(* IEC 61131-3 sources: Test002/ConveyorBelt/Class/SafetyBaseFSoE (part 4) *)

    // if searched path has been found, we already got this pdo in our list
    if (PdoCfg.SourcePathLen = pHelp^.PdoInfo.SourcePathLen) & (PdoCfg.DestPathLen = pHelp^.PdoInfo.DestPathLen) &
      (PdoCfg.InterfaceCRC = pHelp^.PdoInfo.InterfaceCRC) &
      (ToStdLib.MemCmp(dest:= PdoCfg.pSourcePath, source:= pHelp^.PdoInfo.pSourcePath , size:= PdoCfg.SourcePathLen) = 0) &
      (ToStdLib.MemCmp(dest:= PdoCfg.pDestPath,   source:= pHelp^.PdoInfo.pDestPath   , size:= PdoCfg.DestPathLen  ) = 0) then
      // already in buffer => leave function
      return;
    else
      pHelp^.pNext$pvoid := ToStdLib.Malloc(size:=sizeof(t_PdoListElem));
      pHelp := pHelp^.pNext;
    end_if;
  end_if;

  if pHelp <> NIL then
    // allocate memory for the module source path
    pHelp^.PdoInfo.pSourcePath$pVoid := ToStdLib.Malloc(size:=PdoCfg.SourcePathLen);
    if pHelp^.PdoInfo.pSourcePath = NIL then
      SetSafetyState(NewState:=_MemAllocFailed);
      retcode := -1;
      return;
    end_if;

    _memcpy(ptr1:=pHelp^.PdoInfo.pSourcePath, ptr2:=PdoCfg.pSourcePath, cntr:=PdoCfg.SourcePathLen);

    // allocate memory for the module source path
    pHelp^.PdoInfo.pDestPath$pVoid := ToStdLib.Malloc(size:=PdoCfg.DestPathLen);
    if pHelp^.PdoInfo.pDestPath = NIL then
      SetSafetyState(NewState:=_MemAllocFailed);
      retcode := -1;
      return;
    end_if;

    _memcpy(ptr1:=pHelp^.PdoInfo.pDestPath, ptr2:=PdoCfg.pDestPath, cntr:=PdoCfg.DestPathLen);

    pHelp^.PdoInfo.Info           := PdoCfg.Info;
    pHelp^.PdoInfo.InterfaceCRC   := PdoCfg.InterfaceCRC;
    pHelp^.PdoInfo.SourcePathLen  := PdoCfg.SourcePathLen;
    pHelp^.PdoInfo.DestPathLen    := PdoCfg.DestPathLen;
    // length is only zero for non-interface pdos
    if PdoCfg.Info.IsInterfacePDO = FALSE then
      pHelp^.PdoInfo.PdoLen       := 0;   // the length is determined later in method CreateAndSendCfg
    else
      pHelp^.PdoInfo.PdoLen       := PdoCfg.PdoLen;
    end_if;
    pHelp^.PdoInfo.PDO_ID         := 255; // the ID is assigned later by the safety manager of the master domain
    pHelp^.pNext                  := NIL;

    PdoCfgNo += 1;
  else
    SetSafetyState(NewState:=_MemAllocFailed);
    retcode := -1;
    return;
  end_if;

END_FUNCTION

FUNCTION VIRTUAL SafetyBaseFSoE::AddSlaveToCfg
  VAR_INPUT
    pModule 	: ^SafetyBaseFSoE::PathInfoType;
    b_IsOptional 	: BOOL;
    b_IsInterface 	: BOOL;(* := FALSE *)
    InterfaceCRC 	: HDINT;(* := 0 *)
  END_VAR
  VAR
    pHelp : ^t_SlaveListElem;
  END_VAR

  if pFirstSlaveCfg = NIL then
    pFirstSlaveCfg$pVoid := ToStdLib.Malloc(size:=sizeof(t_SlaveListElem));
    pHelp := pFirstSlaveCfg;
  else
    pHelp := pFirstSlaveCfg;
    while pHelp^.pNext <> NIL do
      //if searched path is found, we already got this module in our list
      if (pModule^.ui_PathCompLen = pHelp^.SlaveInfo.CompPathLen) &
        (ToStdLib.MemCmp(dest:= pModule^.p_us_PathComp, source:= pHelp^.SlaveInfo.pCompPath , size:= pModule^.ui_PathCompLen) = 0) then
        // already in buffer => leave function
        return;
      else
        pHelp := pHelp^.pNext;
      end_if;
    end_while;

    //if searched path is found, we already got this module in our list
    if (pModule^.ui_PathCompLen = pHelp^.SlaveInfo.CompPathLen) &
      (ToStdLib.MemCmp(dest:= pModule^.p_us_PathComp, source:= pHelp^.SlaveInfo.pCompPath , size:= pModule^.ui_PathCompLen) = 0) then
      // already in buffer => leave function
      return;
    end_if;

    pHelp^.pNext$pvoid := ToStdLib.Malloc(size:=sizeof(t_SlaveListElem));
    pHelp := pHelp^.pNext;
  end_if;

  if pHelp <> NIL then
    // allocate memory for the module path
    pHelp^.SlaveInfo.PathLen := pModule^.p_us_Path^$UINT + 2;
    pHelp^.SlaveInfo.pPath$pVoid := ToStdLib.Malloc(size:=pHelp^.SlaveInfo.PathLen);
    if pHelp^.SlaveInfo.pPath = NIL then
      SetSafetyState(NewState:=_MemAllocFailed);
      LogError("@0243 (SafetyBaseFSoE::AddSlaveToCfg) Error: Failed to allocate memory for the module path.");
      return;
    end_if;

    _memcpy(ptr1:=pHelp^.SlaveInfo.pPath, ptr2:=pModule^.p_us_Path, cntr:=pHelp^.SlaveInfo.PathLen);

    // allocate memory for the module path
    pHelp^.SlaveInfo.CompPathLen := pModule^.ui_PathCompLen;
    pHelp^.SlaveInfo.pCompPath$pVoid := ToStdLib.Malloc(size:=pHelp^.SlaveInfo.CompPathLen);
    if pHelp^.SlaveInfo.pCompPath = NIL then
      SetSafetyState(NewState:=_MemAllocFailed);
      LogError("@0244 (SafetyBaseFSoE::AddSlaveToCfg) Error: Failed to allocate memory for the compressed module path.");
      return;
    end_if;

    _memcpy(ptr1:=pHelp^.SlaveInfo.pCompPath, ptr2:=pModule^.p_us_PathComp, cntr:=pHelp^.SlaveInfo.CompPathLen);

    pHelp^.SlaveInfo.Info             := 0;
    pHelp^.SlaveInfo.Info.IsOptional  := b_IsOptional;
    pHelp^.SlaveInfo.Info.IsInterface := b_IsInterface;

    pHelp^.SlaveInfo.InterfaceCRC := InterfaceCRC;

    pHelp^.pNext                  := NIL;

    SlaveCfgNo += 1;
  else
    SetSafetyState(NewState:=_MemAllocFailed);
    LogError("@0243 (SafetyBaseFSoE::AddSlaveToCfg) Error: Failed to allocate memory for the new list-element.");
    return;
  end_if;

END_FUNCTION

FUNCTION VIRTUAL SafetyBaseFSoE::FreeCfgLists
  VAR
    pHelpModule : ^t_ModuleListElem;
    pHelpPdo : ^t_PdoListElem;
    pHelpSlave : ^t_SlaveListElem;
//    pHelpUnsafeVar : ^t_UnsafeVarListElem;
  END_VAR

  // while we got module cfgs
  while pFirstModuleCfg do
    pHelpModule := pFirstModuleCfg;
    pFirstModuleCfg := pFirstModuleCfg^.pNext;

    if pHelpModule^.ModuleInfo.pDestCRCs then
      ToStdLib.Free(pHelpModule^.ModuleInfo.pDestCRCs);
    end_if;
    ToStdLib.Free(pHelpModule^.ModuleInfo.pPath);
    ToStdLib.Free(pHelpModule^.ModuleInfo.pCompPath);
    ToStdLib.Free(pHelpModule);
  end_while;
  pFirstModuleCfg := NIL;
  ModuleCfgNo := 0;

  // while we got pdo cfgs
  while pFirstPdoCfg do
    pHelpPdo := pFirstPdoCfg;
    pFirstPdoCfg := pFirstPdoCfg^.pNext;

    ToStdLib.Free(pHelpPdo^.PdoInfo.pSourcePath);
    ToStdLib.Free(pHelpPdo^.PdoInfo.pDestPath);
    ToStdLib.Free(pHelpPdo);
  end_while;
  pFirstPdoCfg := NIL;
  PdoCfgNo := 0;

  // while we got slave cfgs
  while pFirstSlaveCfg do
    pHelpSlave := pFirstSlaveCfg;
    pFirstSlaveCfg := pFirstSlaveCfg^.pNext;

    ToStdLib.Free(pHelpSlave^.SlaveInfo.pPath);
    ToStdLib.Free(pHelpSlave^.SlaveInfo.pCompPath);
    ToStdLib.Free(pHelpSlave);
  end_while;
  pFirstSlaveCfg := NIL;
  SlaveCfgNo := 0;

  FreeFSoEConnectionInfos();

// memory is freed by safety manager
//  // while we got unsafevar cfgs
//  while pFirstUnsafeCfg do
//    pHelpUnsafeVar := pFirstUnsafeCfg;
//    pFirstUnsafeCfg := pFirstUnsafeCfg^.pNext;
//
//    ToStdLib.Free(pHelpUnsafeVar^.UnsafeVarInfo.pName);
//    ToStdLib.Free(pHelpUnsafeVar);
//  end_while;
//  pFirstUnsafeCfg := NIL;
//  UnsafeCfgNo := 0;

  // reduze size of config mem used to 4 (only safety number of cpu module)
  ConfigMemSizeUsed := 4;

END_FUNCTION

FUNCTION VIRTUAL SafetyBaseFSoE::CreateAndSendCfg
  VAR
    pHelpModule       : ^t_ModuleListElem;
    pHelpPdo          : ^t_PdoListElem;
    pHelpSlave        : ^t_SlaveListElem;
    pHelpConnection   : ^t_FSoEConnectionDetails;
    pCfg              : ^void;
    TmpPathLen        : UINT;
    MyPara 	          : CmdStruct;
    MyResult	        : results;
    AddConfigSize     : UDINT;
    i                 : UDINT;
  END_VAR

(*
    Memory structure:
      4 Byte: SafetyNumber of CPU (is already there from initialisation in CSCP011_IM::InitSafeModule)
      1 Byte: Number of module configurations which are following
      for every module configuration (first is always the CPU itself)
        1 Byte: Info
        4 Byte: Interface Frame Source SafetyNumber (0 if it is no source for interface frames)
        4 Byte: Interface Frame CRC
        1 Byte: Number of destination inferface frame CRCs
        x Byte: Destination interface frame CRCs (number * sizeof(HDINT)
        2 Byte: Length of hardware path
        x Byte (depending on length in the 2 byte before): Hardwarepath
        2 Byte: Length of compressed hardware path
        x Byte (depending on length in the 2 byte before): Compressed Hardwarepath
        1 Byte: PDO out length for this module
      1 Byte: Number of pdo configurations which are following
      for every PDO configuration
        1 Byte: PDO length
        1 Byte: Interface frame info
        4 Byte: Interface CRC
        2 Byte: Length of source hardware path
        x Byte (depending on length in the 2 byte before): Hardwarepath of source
        2 Byte: Length of destination hardware path
        x Byte (depending on length in the 2 byte before): Hardwarepath of destination
      1 Byte: Number of slave configurations which are following
      for every slave configuration
        1 Byte: Info
        4 Byte: InterfaceCRC
        2 Byte: Length of hardware path
        x Byte (depending on length in the 2 byte before): Hardwarepath
        2 Byte: Length of compressed hardware path
        x Byte (depending on length in the 2 byte before): Compressed Hardwarepath
      2 Byte: Number of connection infos which are following
      for every FSoE connection info
        2 Byte: ConnectionID
        1 Byte: ConnectionState
        1 Byte: Flags // Actually, type is 4 bytes in size but for compatibility reasons it is still used as 1 byte. As a result, bits 9-32 are currently not used.
        4 Byte: Master safety number

only if feature available:
        2 Byte: Transmission time in ms

        2 Byte: Offset where to read from master
        2 Byte: Size of data to read from master (and write to slave)
        2 Byte: Offset where to write to master
        2 Byte: Size of data to write to master (and read from slave)
        2 Byte: SlaveAddress
        2 Byte: Length of slave hardware path
        x Byte (depending on length in the 2 byte before): Slave hardware path
        2 Byte: Length of compressed slave hardware path
        x Byte (depending on length in the 2 byte before): Compressed slave hardware path
        2 Byte: Offset where to read from slave
        2 Byte: Offset where to write to slave
*)

  // check if there is memory and if the only thing inside is the safety number
  if pConfigMem & (ConfigMemSizeUsed = 4) then
    // insert the safety number
    pConfigMem^$UDINT := SafetyNumber;

    // pCfg points to the next memory we have to write to => set it to the memory after the safety number
    pCfg := pConfigMem + ConfigMemSizeUsed;

    // add all module configurations to memory
    if pFirstModuleCfg then
      // add number of module configurations to memory (no need to check the memory here, because already 512 bytes are allocated)
      pCfg^$USINT       := ModuleCfgNo;
      pCfg              += sizeof(USINT);
      ConfigMemSizeUsed += sizeof(USINT);

      pHelpModule := pFirstModuleCfg;
      // go through list
      while pHelpModule do
        // add the elements

        // check if we have enough memory to add the next module
        AddConfigSize := sizeof(BSINT) + sizeof(HDINT) + sizeof(HDINT) + sizeof(UINT) + pHelpModule^.ModuleInfo.PathLen + sizeof(UINT) + pHelpModule^.ModuleInfo.CompPathLen + sizeof(USINT);
        if pHelpModule^.ModuleInfo.Info.IsInterfaceDest then
          AddConfigSize += sizeof(USINT) + pHelpModule^.ModuleInfo.DestCRCNo * sizeof(HDINT);
        end_if;

        pCfg := CheckConfigMemSize(AddConfigSize);
        if pCfg = NIL then
          // error message already logged by function
          return;
        end_if;

        // info
        pCfg^$BSINT := pHelpModule^.ModuleInfo.Info;
        pCfg              += sizeof(BSINT);
        ConfigMemSizeUsed += sizeof(BSINT);

        // safety number of interface frame source (if it is one)
        pCfg^$HDINT := pHelpModule^.ModuleInfo.SafetyNbr;
        pCfg              += sizeof(HDINT);
        ConfigMemSizeUsed += sizeof(HDINT);

        // interface CRC of interface frame
        pCfg^$HDINT := pHelpModule^.ModuleInfo.InterfaceCRC;
        pCfg              += sizeof(HDINT);
        ConfigMemSizeUsed += sizeof(HDINT);

        // if its also interface frame destination send the corresponding interface CRCs
        if pHelpModule^.ModuleInfo.Info.IsInterfaceDest then
          TmpPathLen := pHelpModule^.ModuleInfo.DestCRCNo; // save some time with this local variable
          pCfg^$USINT := TmpPathLen$USINT;
          pCfg              += sizeof(USINT);
          ConfigMemSizeUsed += sizeof(USINT);

          _memcpy(ptr1:=pCfg, ptr2:=pHelpModule^.ModuleInfo.pDestCRCs, cntr:=TmpPathLen * sizeof(HDINT));
          pCfg += TmpPathLen * sizeof(HDINT);
          ConfigMemSizeUsed += TmpPathLen * sizeof(HDINT);
        end_if;

        // uncompressed module path
        TmpPathLen := pHelpModule^.ModuleInfo.PathLen; // save some time with this local variable
        pCfg^$UINT := TmpPathLen;
        pCfg              += sizeof(UINT);
        ConfigMemSizeUsed += sizeof(UINT);

        _memcpy(ptr1:=pCfg, ptr2:=pHelpModule^.ModuleInfo.pPath, cntr:=TmpPathLen);
        pCfg += TmpPathLen;
        ConfigMemSizeUsed += TmpPathLen;

        // compressed module path
        TmpPathLen := pHelpModule^.ModuleInfo.CompPathLen; // save some time with this local variable
        pCfg^$UINT := TmpPathLen;
        pCfg              += sizeof(UINT);
        ConfigMemSizeUsed += sizeof(UINT);

        _memcpy(ptr1:=pCfg, ptr2:=pHelpModule^.ModuleInfo.pCompPath, cntr:=TmpPathLen);
        pCfg += TmpPathLen;
        ConfigMemSizeUsed += TmpPathLen;

        // PDO out length for this module (to assign the length to the pdo configurations)
        pCfg^$USINT := pHelpModule^.ModuleInfo.PdoOutLen;
        pCfg              += sizeof(USINT);
        ConfigMemSizeUsed += sizeof(USINT);

        pHelpModule := pHelpModule^.pNext;
      end_while;

      pCfg := CheckConfigMemSize(sizeof(USINT));
      if pCfg = NIL then
        // error message already logged by function
        return;
      end_if;

      // add number of pdo configurations to memory
      pCfg^$USINT := PdoCfgNo;
      pCfg              += sizeof(USINT);
      ConfigMemSizeUsed += sizeof(USINT);

      // add all pdo configurations to memory (module configs must be available, to find out the PDO length)
      if pFirstPdoCfg then
        pHelpPdo := pFirstPdoCfg;
        // go through list
        while pHelpPdo do
          // add the elements

          // check if we have enough memory to add the next module
          AddConfigSize := sizeof(USINT) + sizeof(BSINT) + sizeof(HDINT) + sizeof(UINT) + pHelpPdo^.PdoInfo.SourcePathLen + sizeof(UINT) + pHelpPdo^.PdoInfo.DestPathLen;
          pCfg := CheckConfigMemSize(AddConfigSize);
          if pCfg = NIL then
            // error message already logged by function
            return;
          end_if;

          // first of all we have to find out the pdo length of this element => search the module configurations until we find our source and copy the pdo length
          if pHelpPdo^.PdoInfo.PdoLen = 0 then
            pHelpModule := pFirstModuleCfg;
            // go through list
            while pHelpModule do
              // if the path of the source module matches, save the pdolength of this module
              if (pHelpPdo^.PdoInfo.SourcePathLen = pHelpModule^.ModuleInfo.PathLen) & (ToStdLib.MemCmp(dest:= pHelpPdo^.PdoInfo.pSourcePath, source:= pHelpModule^.ModuleInfo.pPath , size:= pHelpPdo^.PdoInfo.SourcePathLen) = 0) then
                pHelpPdo^.PdoInfo.PdoLen := pHelpModule^.ModuleInfo.PdoOutLen;
                exit;
              end_if;
              pHelpModule := pHelpModule^.pNext;
            end_while;
          end_if;

          // PDO Length
          pCfg^$USINT := pHelpPdo^.PdoInfo.PdoLen;
          pCfg              += sizeof(USINT);
          ConfigMemSizeUsed += sizeof(USINT);

          // info
          pCfg^$BSINT := pHelpPdo^.PdoInfo.Info;
          pCfg              += sizeof(BSINT);
          ConfigMemSizeUsed += sizeof(BSINT);

          // interface CRC
          pCfg^$HDINT := pHelpPdo^.PdoInfo.InterfaceCRC;
          pCfg              += sizeof(HDINT);
          ConfigMemSizeUsed += sizeof(HDINT);

          // Source Path Length
          TmpPathLen := pHelpPdo^.PdoInfo.SourcePathLen; // save some time with this local variable
          pCfg^$UINT := TmpPathLen;
          pCfg              += sizeof(UINT);
          ConfigMemSizeUsed += sizeof(UINT);

          // Source Path
          _memcpy(ptr1:=pCfg, ptr2:=pHelpPdo^.PdoInfo.pSourcePath, cntr:=TmpPathLen);
          pCfg += TmpPathLen;
          ConfigMemSizeUsed += TmpPathLen;

          // Destination Path Length
          TmpPathLen := pHelpPdo^.PdoInfo.DestPathLen; // save some time with this local variable
          pCfg^$UINT := TmpPathLen;
          pCfg              += sizeof(UINT);
          ConfigMemSizeUsed += sizeof(UINT);

          // Destination Path
          _memcpy(ptr1:=pCfg, ptr2:=pHelpPdo^.PdoInfo.pDestPath, cntr:=TmpPathLen);
          pCfg += TmpPathLen;
          ConfigMemSizeUsed += TmpPathLen;

          pHelpPdo := pHelpPdo^.pNext;
        end_while;
      end_if;

      pCfg := CheckConfigMemSize(sizeof(USINT));
      if pCfg = NIL then
        // error message already logged by function
        return;
      end_if;

      // add number of slave configurations to memory
      pCfg^$USINT       := SlaveCfgNo;
      pCfg              += sizeof(USINT);
      ConfigMemSizeUsed += sizeof(USINT);

      pHelpSlave := pFirstSlaveCfg;
      // go through list
      while pHelpSlave do
        // add the elements

        // check if we have enough memory to add the next module
        AddConfigSize := sizeof(BSINT) + sizeof(HDINT) + sizeof(UINT) + pHelpSlave^.SlaveInfo.PathLen + sizeof(UINT) + pHelpSlave^.SlaveInfo.CompPathLen;

        pCfg := CheckConfigMemSize(AddConfigSize);
        if pCfg = NIL then
          // error message already logged by function
          return;
        end_if;

        // info
        pCfg^$BSINT := pHelpSlave^.SlaveInfo.Info;
        pCfg              += sizeof(BSINT);
        ConfigMemSizeUsed += sizeof(BSINT);

        // InterfaceCRC
        pCfg^$HDINT := pHelpSlave^.SlaveInfo.InterfaceCRC;
        pCfg              += sizeof(HDINT);
        ConfigMemSizeUsed += sizeof(HDINT);

        // uncompressed Slave path
        TmpPathLen := pHelpSlave^.SlaveInfo.PathLen; // save some time with this local variable
        pCfg^$UINT := TmpPathLen;
        pCfg              += sizeof(UINT);
        ConfigMemSizeUsed += sizeof(UINT);

        _memcpy(ptr1:=pCfg, ptr2:=pHelpSlave^.SlaveInfo.pPath, cntr:=TmpPathLen);
        pCfg += TmpPathLen;
        ConfigMemSizeUsed += TmpPathLen;

        // compressed Slave path
        TmpPathLen := pHelpSlave^.SlaveInfo.CompPathLen; // save some time with this local variable
        pCfg^$UINT := TmpPathLen;
        pCfg              += sizeof(UINT);
        ConfigMemSizeUsed += sizeof(UINT);

        _memcpy(ptr1:=pCfg, ptr2:=pHelpSlave^.SlaveInfo.pCompPath, cntr:=TmpPathLen);
        pCfg += TmpPathLen;
        ConfigMemSizeUsed += TmpPathLen;

        pHelpSlave := pHelpSlave^.pNext;
      end_while;

    else
      // add number of module, pdo and slave configurations to memory (all as 0)

      pCfg := CheckConfigMemSize(3*sizeof(USINT));
      if pCfg = NIL then
        // error message already logged by function
        return;
      end_if;

      // no module configs
      pCfg^$USINT := 0;
      pCfg              += sizeof(USINT);
      ConfigMemSizeUsed += sizeof(USINT);

      // no pdo configs
      pCfg^$USINT := 0;
      pCfg              += sizeof(USINT);
      ConfigMemSizeUsed += sizeof(USINT);

      // no slave configs
      pCfg^$USINT := 0;
      pCfg              += sizeof(USINT);
      ConfigMemSizeUsed += sizeof(USINT);
    end_if;

    pCfg := CheckConfigMemSize(sizeof(UINT));
    if pCfg = NIL then
      // error message already logged by function
      return;
    end_if;

    // number of connection details
    pCfg^$UINT := ConnectionInfos.ConnectionNo$UINT;
    pCfg              += sizeof(UINT);
    ConfigMemSizeUsed += sizeof(UINT);

    if ConnectionInfos.ConnectionNo then

      pHelpConnection := ConnectionInfos.pFirstConnection;
      for i := 0 to (ConnectionInfos.ConnectionNo-1) do
        // add the elements

        // check if we have enough memory to add the next connection
        AddConfigSize := sizeof(UINT) + sizeof(USINT) + sizeof(USINT) + bdFeatureEnable.FSoEFlags_4ByteSize * 3 * sizeof(USINT) + sizeof(HDINT) +
                         6 * sizeof(UINT) + pHelpConnection^.SlavePathLen + sizeof(UINT) + pHelpConnection^.SlavePathCompLen + 2 * sizeof(UINT);

        if bdFeatureEnable.TransmissionTimeInConfig then
          AddConfigSize += sizeof(UINT);
        end_if;

        pCfg := CheckConfigMemSize(AddConfigSize);
        if pCfg = NIL then
          // error message already logged by function
          return;
        end_if;

        // connection ID
        pCfg^$UINT        := pHelpConnection^.ConnectionID;
        pCfg              += sizeof(UINT);
        ConfigMemSizeUsed += sizeof(UINT);

        // connection state
        pCfg^$USINT       := pHelpConnection^.ConnectionState$USINT;
        pCfg              += sizeof(USINT);
        ConfigMemSizeUsed += sizeof(USINT);

        // flags
        // In older Safety manager versions this flag is only used as 1 byte. Now we use 4 byte if safetymanager supports this
        if bdFeatureEnable.FSoEFlags_4ByteSize then
          pCfg^$t_FSoEFlags := pHelpConnection^.Flags;
          pCfg              += sizeof(t_FSoEFlags);
          ConfigMemSizeUsed += sizeof(t_FSoEFlags);
        else
          pCfg^$USINT       := pHelpConnection^.Flags$USINT;
          pCfg              += sizeof(USINT);
          ConfigMemSizeUsed += sizeof(USINT);
        end_if;

        // master safety number
        pCfg^$HDINT       := pHelpConnection^.OwnerSafetyNbr;
        pCfg              += sizeof(HDINT);
        ConfigMemSizeUsed += sizeof(HDINT);

        // the feature is not available in older safety manager classes, so we have to do this for compatibility reasons
        if bdFeatureEnable.TransmissionTimeInConfig then
          // transmission time settings from safety designer
          pCfg^$UINT        := pHelpConnection^.TransmissionTime_ms;
          pCfg              += sizeof(UINT);
          ConfigMemSizeUsed += sizeof(UINT);
        end_if;

        // offset where to read from master
        pCfg^$UINT        := pHelpConnection^.MasterReadOffset;
        pCfg              += sizeof(UINT);
        ConfigMemSizeUsed += sizeof(UINT);

        // size of data to read from master (and write to slave)
        pCfg^$UINT        := pHelpConnection^.MasterReadSize;
        pCfg              += sizeof(UINT);
        ConfigMemSizeUsed += sizeof(UINT);

        // offset where to write to master
        pCfg^$UINT        := pHelpConnection^.MasterWriteOffset;
        pCfg              += sizeof(UINT);
        ConfigMemSizeUsed += sizeof(UINT);

        // size of data to write to master (and read from slave)
        pCfg^$UINT        := pHelpConnection^.MasterWriteSize;
        pCfg              += sizeof(UINT);
        ConfigMemSizeUsed += sizeof(UINT);

        // slave address
        pCfg^$UINT        := pHelpConnection^.SlaveAddress;
        pCfg              += sizeof(UINT);
        ConfigMemSizeUsed += sizeof(UINT);

        // uncompressed slave path
        TmpPathLen        := pHelpConnection^.SlavePathLen; // save some time with this local variable
        pCfg^$UINT        := TmpPathLen;
        pCfg              += sizeof(UINT);
        ConfigMemSizeUsed += sizeof(UINT);

        _memcpy(ptr1:=pCfg, ptr2:=pHelpConnection^.pSlavePath, cntr:=TmpPathLen);
        pCfg              += TmpPathLen;
        ConfigMemSizeUsed += TmpPathLen;

        // compressed slave path
        TmpPathLen        := pHelpConnection^.SlavePathCompLen; // save some time with this local variable
        pCfg^$UINT        := TmpPathLen;
        pCfg              += sizeof(UINT);
        ConfigMemSizeUsed += sizeof(UINT);

        _memcpy(ptr1:=pCfg, ptr2:=pHelpConnection^.pSlavePathComp, cntr:=TmpPathLen);
        pCfg              += TmpPathLen;
        ConfigMemSizeUsed += TmpPathLen;

        // offset where to read from slave
        pCfg^$UINT        := pHelpConnection^.SlaveReadOffset;
        pCfg              += sizeof(UINT);
        ConfigMemSizeUsed += sizeof(UINT);

        // offset where to write to slave
        pCfg^$UINT        := pHelpConnection^.SlaveWriteOffset;
        pCfg              += sizeof(UINT);
        ConfigMemSizeUsed += sizeof(UINT);

        pHelpConnection += sizeof(t_FSoEConnectionDetails);
      end_for;
    end_if;

    MyPara.uiCmd := CMD_SM_FSOE_CFG_TO_MANAGER;
    MyPara.aPara[0] := ConfigMemSizeUsed$DINT;
    MyPara.aPara[1] := pConfigMem$DINT;
    if pSafetyManagerThis^.NewInst(#MyPara, #MyResult) = READY then
      // the manager takes care of our memory from now on
      pFirstSlaveCfg := NIL;
    end_if;

    // now tell the manager, what kind of configuration we have
    MyPara.uiCmd := CMD_SM_NEW_CFG_TYPE;
    MyPara.aPara[0] := SafetyNumber$DINT;
    MyPara.aPara[1] := NewConfigType;
    pSafetyManagerThis^.NewInst(#MyPara, #MyResult);
  else
    LogError("@0245 (SafetyBaseFSoE::CreateAndSendCfg) No config memory or invalid memory size usage.");
  end_if;

END_FUNCTION

#pragma warning(disable: 73)
FUNCTION VIRTUAL SafetyBaseFSoE::CheckVariant
  VAR_INPUT
    us_ActVariant 	: USINT;
  END_VAR
  VAR_OUTPUT
    b_IsOK 	: BOOL;
  END_VAR

  // if the overwritten methods are getting deleted, we already have a code for compatiblity here
  b_IsOK := TRUE; // FALSE;

END_FUNCTION
#pragma warning(default: 73)

FUNCTION SafetyBaseFSoE::SendAllUnsafeValues
  VAR
    pHelpUnsafeOut : ^UnsafeIORoutingElement;
  END_VAR

  // mark all unsafe values as not sent
  pHelpUnsafeOut := p_UnsafeInputsTable;
  while pHelpUnsafeOut do
    pHelpUnsafeOut^.b_AlreadyTransmitted := FALSE;

    pHelpUnsafeOut := pHelpUnsafeOut^.pNext;
  end_while;

  // reset the actual pointer
  pUnsafeInElement := NIL;

END_FUNCTION

FUNCTION SafetyBaseFSoE::GetDestinationCRCs
  VAR
    pHelpModule : ^t_ModuleListElem;
    pHelpPdo : ^t_PdoListElem;
  END_VAR

  // go through the module list
  pHelpModule := pFirstModuleCfg;
  while pHelpModule do
    pHelpPdo := pFirstPdoCfg;
    while pHelpPdo do
      // search in the PDOs if this module is an interface frame destination somewhere
      if pHelpPdo^.PdoInfo.Info.IsInterfacePDO then
        if (pHelpPdo^.PdoInfo.DestPathLen = pHelpModule^.ModuleInfo.PathLen) &
         (ToStdLib.MemCmp(dest:= pHelpModule^.ModuleInfo.pPath, source:= pHelpPdo^.PdoInfo.pDestPath , size:= pHelpModule^.ModuleInfo.PathLen) = 0) then
          pHelpModule^.ModuleInfo.Info.IsInterfaceDest := TRUE;
          if pHelpModule^.ModuleInfo.DestCRCNo & pHelpModule^.ModuleInfo.pDestCRCs then
            pHelpModule^.ModuleInfo.pDestCRCs$^void := ToStdLib.ReAlloc(mptr:=pHelpModule^.ModuleInfo.pDestCRCs, newsize:=(pHelpModule^.ModuleInfo.DestCRCNo+1) * sizeof(HDINT));
          else
            pHelpModule^.ModuleInfo.pDestCRCs$^void := ToStdLib.Malloc(sizeof(HDINT));
          end_if;

          (pHelpModule^.ModuleInfo.pDestCRCs + pHelpModule^.ModuleInfo.DestCRCNo * sizeof(HDINT))^ := pHelpPdo^.PdoInfo.InterfaceCRC;

          pHelpModule^.ModuleInfo.DestCRCNo += 1;
        end_if;
      else
        // if this is module is optional and it's the source of the PDO => the pdo is also optional
        if pHelpModule^.ModuleInfo.Info.IsOptional & (pHelpPdo^.PdoInfo.SourcePathLen = pHelpModule^.ModuleInfo.PathLen) &
         (ToStdLib.MemCmp(dest:= pHelpModule^.ModuleInfo.pPath, source:= pHelpPdo^.PdoInfo.pSourcePath , size:= pHelpModule^.ModuleInfo.PathLen) = 0) then
          pHelpPdo^.PdoInfo.Info.IsOptional := TRUE;
        end_if;
      end_if;

      pHelpPdo := pHelpPdo^.pNext;
    end_while;

    pHelpModule := pHelpModule^.pNext;
  end_while;

END_FUNCTION

FUNCTION SafetyBaseFSoE::CountBits
  VAR_INPUT
    BitMask 	: BDINT;
  END_VAR
  VAR_OUTPUT
    BitNo 	: UDINT;
  END_VAR

  BitNo := 0;

  while BitMask do
    BitMask := BitMask AND (BitMask - 1);
    BitNo += 1;
  end_while;

END_FUNCTION

FUNCTION VIRTUAL SafetyBaseFSoE::IsOptimizedCPU
  VAR_OUTPUT
    IsOptimized 	: DINT;
  END_VAR

  // every derivation of this class is an optimized cpu, which means the SBF_SDO_COMMAND_WRITE_VALUES command is available to save time in communication of unsafe variables
  IsOptimized := TRUE;

END_FUNCTION

FUNCTION VIRTUAL SafetyBaseFSoE::CheckConfigMemSize
  VAR_INPUT
    AddConfigSize 	: UDINT;
  END_VAR
  VAR_OUTPUT
    pCfg 	: ^void;
  END_VAR
  VAR
    pTempMem  : ^void;
  END_VAR

  pCfg := NIL;

  if ((ConfigMemSizeUsed + AddConfigSize) > ConfigMemSize) then
    // if there isn't enough memory => reallocate
    pTempMem := ToStdLib.ReAlloc(mptr:=pConfigMem, newsize:=GetNewMemSize(ConfigMemSizeUsed + AddConfigSize));
    IF pTempMem <> NIL THEN
      pConfigMem := pTempMem;
      ConfigMemSize := GetNewMemSize(ConfigMemSizeUsed + AddConfigSize);
    ELSE
      SetSafetyState(NewState:=_MemAllocFailed);
      LogError("@0246 (SafetyBaseFSoE::CreateAndSendCfg) Failed to reallocate configuration memory!");
      return;
    END_IF;
  end_if;

  pCfg := pConfigMem + ConfigMemSizeUsed;

END_FUNCTION

FUNCTION SafetyBaseFSoE::DToH
  VAR_INPUT
    pt 	: ^CHAR;
    value 	: DINT;
  END_VAR
  VAR
    val  : UDINT;
  END_VAR

  // this method converts a single byte into a zero-terminated hexstring like 0xA4 => "A4"
  val := value$UDINT;

  // zero termination
  (pt + 2)^ := 0;

  // start with the low nibble
  if (val AND 16#F) < 10 then
    (pt + 1)^ := (val AND 16#F)$USINT + '0';
  else
    (pt + 1)^ := (val AND 16#F)$USINT - 10 + 'A';
  end_if;

  // now get the high nibble
  val := val / 16;

  if (val AND 16#F) < 10 then
    pt^ := (val AND 16#F)$USINT + '0';
  else
    pt^ := (val AND 16#F)$USINT - 10 + 'A';
  end_if;

END_FUNCTION

FUNCTION SafetyBaseFSoE::LogHWPath
  VAR_INPUT
    pString 	: ^CHAR;
    pHWPath 	: ^USINT;
  END_VAR
  VAR
    TempStr       : ARRAY [0..99] OF CHAR;
    TraceVal      : USINT;
    i             : UINT;
    MyMsg         : ARRAY [0..599] OF CHAR;
  END_VAR

  if pString & pHWPath then

    _strncpy(dest:=#MyMsg[0], src:=pString, max:=200);

    TraceVal := pHWPath^;
    if TraceVal then
      TraceVal += 2; //show also the length
      i := 0;
      while (TraceVal >= 1) & (i < 95) do
        DToH(#TempStr[i], pHWPath^$USINT);
        i += 2; // 2 chars per byte
        TempStr[i] := ' ';
        i += 1;
        pHWPath += 1;
        TraceVal -= 1;
      end_while;
      TempStr[i] := 0;

      _strcat( dest:=#MyMsg[0], src:=#TempStr[0]);
    end_if;

#ifdef HWC_LogError
    HWC_LogError(this, #MyMsg[0]);
#endif
  end_if;

END_FUNCTION

FUNCTION VIRTUAL GLOBAL SafetyBaseFSoE::QuitComError::Write
  VAR_INPUT
    input (EAX) 	: DINT;
  END_VAR
  VAR_OUTPUT
    result (EAX) 	: DINT;
  END_VAR

  result := input;

  if ErrorState then
    if b_QuitErrorAvailable then
      // remember to do it in next background
      QuitComError := 2;
    else
      // remember. that there has been a manual quit (for writing PDOs in PostScan)
      b_ManualQuit := TRUE;

      // remember to do it in next cyclic
      QuitComError := 1;
    end_if;
  end_if;

  // refresh the server on the outer object
  RefreshAsySrv();

END_FUNCTION

FUNCTION VIRTUAL GLOBAL SafetyBaseFSoE::ClassSvr::NewInst
  VAR_INPUT
    pPara 	: ^CmdStruct;
    pResult 	: ^results;
  END_VAR
  VAR_OUTPUT
    ret_code 	: iprStates;
  END_VAR
  VAR
    OldClassState : SafetyConfigStateType;
    pPDOInputBuffer : ^PDOInputBuffer;
    i, j : UINT;
    Found : BOOL;
    sd_retval : DINT;
    GetStateResp   : GetStateResponseType;
  END_VAR

  ret_code := READY;

  CASE pPara^.uiCmd OF
//**********************************************************************************************************************************************************
    CMD_SM_INIT_FINISHED:
      // the safety manager has finished his administration work (e.g. connecting the domains)
      b_ManagerInitialisationFinished := TRUE;

      // optional modules may not be available
      ud_OptionalTimeoutStart := ops.tAbsolute;

//**********************************************************************************************************************************************************
    CMD_SM_FIRST_CONNECT_READY:
      // the safety manager has finished first time connecting the domains
      b_ManagerReadyForSDO := TRUE;

//**********************************************************************************************************************************************************
    CMD_SM_DISCONNECT:
      b_ManagerInitialisationFinished := FALSE;
      b_ManagerReadyForSDO := FALSE;

      // wait again to send bus ready signal
      if SafetyState <> _ReinitConfig then
        SetSafetyState(NewState:=_WaitForSynchronicity);
      end_if;
      UnsafeScheduler := UnsafeSchedulerSetBusReady;
      us_SetBusReadyState := WaitPDOsSyncron;

//**********************************************************************************************************************************************************
    CMD_SM_SDO_TO_MODULE:
#ifdef DO_DEBUG
      DOCheck(pFrame:=(pPara^.aPara[1])$^t_SDOStdHeader, pCheckStruct:=#SDOWrite);
#endif

      AddSDOToBuffer(p_us_Message := pPara^.aPara[1]$^USINT, us_length := pPara^.aPara[0]$USINT);

//**********************************************************************************************************************************************************
    CMD_SM_GET_SAFETY_NUMBER:
      // check if pointer is valid
      if pPara^.aPara[0] then
        ((pPara^.aPara[0])$^UDINT)^ := SafetyNumber;
      end_if;
//**********************************************************************************************************************************************************
    CMD_SM_ADD_INPUT_PDO:
      // check if the information if it's an interface frame (stored at pPara^.aPara[9]$BOOL) is valid
      if pPara^.aPara[8]$HDINT = SM_IF_VALIDITY_MARK then
        sd_retval :=
        AddPDOToInputBuffer(ud_p2Buffer         := pPara^.aPara[0]$UDINT
                          , ud_SafetyNr         := pPara^.aPara[2]$UDINT
                          , b_IsOptional        := pPara^.aPara[4]$BOOL
                          , ui_PdoLen           := pPara^.aPara[3]$UINT
                          , ui_TargetOffset     := pPara^.aPara[7]$UINT
                          , b_IsInterfaceFrame  := pPara^.aPara[9]$BOOL
                          );
      else
        sd_retval :=
        AddPDOToInputBuffer(ud_p2Buffer         := pPara^.aPara[0]$UDINT
                          , ud_SafetyNr         := pPara^.aPara[2]$UDINT
                          , b_IsOptional        := pPara^.aPara[4]$BOOL
                          , ui_PdoLen           := pPara^.aPara[3]$UINT
                          , ui_TargetOffset     := pPara^.aPara[7]$UINT
                          );
      end_if;

      if sd_retval then
        ret_code := ERROR;
      end_if;

//**********************************************************************************************************************************************************
    CMD_SM_ADD_OUTPUT_PDO:
      // if it's an interface frame, we return the pointer to the second PDO frame which is the interface pdo frame
//      if pPara^.aPara[0] = 1 then
//        // skip the first PDO
//        pResult^.aData[0]$UDINT := GetPointer2IFPDOBuffer();    // pointer to local memory
//        pResult^.aData[4]$UDINT := ud_LocalMoveIFSourceAddr;    // pointer to DPRAM
//        pResult^.aData[8]$UDINT := ud_LocalIFReadHandle;        // handle for varan access
//        pResult^.aData[12]$UDINT:= ud_LocalIFReadOffset;        // offset inside the varan data
//      else
//        // otherwise just get the pointer to the PDO read data
//        pResult^.aData[0]$UDINT := GetPointer2PDOBuffer();      // pointer to local memory
//        pResult^.aData[4]$UDINT := ud_LocalMoveSourceAddr;      // pointer to DPRAM
//        pResult^.aData[8]$UDINT := ud_LocalReadHandle;          // handle for varan access
//        pResult^.aData[12]$UDINT:= ud_LocalReadOffset;          // offset insid the varan data
//      end_if;

      // return the pointer to the Buffer (is linear local memory, so the offset can be added later)
      pResult^.aData[0]$UDINT := GetPointer2PDOBuffer();
      pResult^.uiLng := 4;

//**********************************************************************************************************************************************************
    CMD_SM_REMOVE_INPUT_PDO:
      // we lost connection to other systems => we have to initialize again! remove old input PDOs

      if ui_cnt_PDOInputBuffer then
        // save the old state of the class and set it temporarily to "module not found" to prevent update rt from crashing
        OldClassState := SafetyState;
        SetSafetyState(NewState:=_ModuleNotFound);

        // search for the PDO
        Found := FALSE;
        pPDOInputBuffer := #aPDOInputBuffer[0];
        for i := 0 to (ui_cnt_PDOInputBuffer-1) do
          if pPDOInputBuffer^.ud_p2Buffer = pPara^.aPara[0]$UDINT then
            Found := TRUE;
            exit;
          end_if;

          pPDOInputBuffer += sizeof(PDOInputBuffer);
        end_for;

        // if we found the PDO => remove it from memory (move the memory behind the found PDO over the place of the found PDO)
        if Found then
          // if it's last entry (no entries have to be moved) => we only have to copy some memory if it's not the last
          if i < (ui_cnt_PDOInputBuffer-1) then
            for j := i to (ui_cnt_PDOInputBuffer-2) do
              aPDOInputBuffer[j] := aPDOInputBuffer[j+1];
            end_for;
          end_if;
          ui_cnt_PDOInputBuffer -= 1;

          if ui_cnt_PDOInputBuffer = 0 then
            if ModuleSyncNo & (SafetyState <> _SafetyClassOK) then
              ModuleSyncNo -= 1;
            end_if;
          end_if;

//        else
//          LogError("@ZZZZ (SafetyBaseFSoE::State::NewInst) CMD_SM_REMOVE_INPUT_PDO failed! Couldn't find specified PDO!");
        end_if;

        // restore old class state
        SetSafetyState(NewState:=OldClassState);
//      else
//        LogError("@ZZZZ (SafetyBaseFSoE::State::NewInst) CMD_SM_REMOVE_INPUT_PDO failed! No input PDOs found!");
      end_if;

//*****************************************************************************
//** COMMANDS FROM BUS INTERFACE                                             **
//*****************************************************************************

//**********************************************************************************************************************************************************
    _BUS_IF_HWCONNECT :
      // device has been connected
      ConnectEvent();
      pResult^.aData[0] := _BUS_IF_RETVAL_OK;

//**********************************************************************************************************************************************************
    _BUS_IF_HWDISCONNECT :
      // device has been disconnected
      DisconnectEvent();
      pResult^.aData[0] := _BUS_IF_RETVAL_OK;

//**********************************************************************************************************************************************************
    _BUS_IF_HWINTERRUPT :
      // error at device which may lead to a disconnect or replace the disconnect callback
      InterruptEvent();
      pResult^.aData[0] := _BUS_IF_RETVAL_OK;

//**********************************************************************************************************************************************************
    _BUS_IF_CHECK_DEVICE_ID :
      // check for correct device id
      pResult^.aData[0] := (DeviceID = pPara^.aPara[0]$UDINT);

//**********************************************************************************************************************************************************
    _BUS_IF_RESET_DETECTED:
      if SafetyState = _SafetyClassOK then
        SafetyState := _LostPowerSupply;
      end_if;

//**********************************************************************************************************************************************************
    _BUS_IF_RESET_GONE_DETECTED:
      if SafetyState = _LostPowerSupply then
        SafetyState := _SafetyClassOK;
      end_if;

//**********************************************************************************************************************************************************

//*****************************************************************************
//** COMMANDS FROM OTHER SAFETYMODULES                                       **
//*****************************************************************************

//**********************************************************************************************************************************************************
    CMD_SM_ADD_SDO_TO_BUFFER:
      sd_retval := AddSDOToBuffer(p_us_message:=pPara^.aPara[0]$^USINT, us_length:=pPara^.aPara[1]$USINT);
      if sd_retval then
        ret_code := ERROR;
      end_if;

      pResult^.aData[0]$DINT := sd_retval;

//**********************************************************************************************************************************************************
    CMD_SM_CONFIG_SAFETY_CPU:
      pResult^.aData[0]$UDINT := ConfigSafetyCpu();

//**********************************************************************************************************************************************************
    CMD_SM_CONFIG_SAFETY_INPUT:
      pResult^.aData[0]$UDINT := ConfigSafetyInput(ud_SafeNrCPU         := pPara^.aPara[0]$HDINT
                                                 , ud_thisp             := pPara^.aPara[1]$UDINT
                                                 , p_PDOBuffer          := pPara^.aPara[2]$^UDINT
                                                 );

//**********************************************************************************************************************************************************
    CMD_SM_CONFIG_SAFETY_OUTPUT:
      pResult^.aData[0]$UDINT := ConfigSafetyOutput(ud_SafeNrCPU        := pPara^.aPara[0]$HDINT
                                                  , ud_thisp            := pPara^.aPara[1]$UDINT
                                                  , ud_p_PDOBuffer      := pPara^.aPara[2]$UDINT
                                                  , pObject             := pPara^.aPara[3]$^PathInfoType
                                                  , b_IsOptional        := pPara^.aPara[6]$BOOL
                                                  );

//**********************************************************************************************************************************************************
    CMD_SM_REMOVE_CPU_FROM_TABLE:
      RemoveCPUFromTable(ud_SafetyNr := pPara^.aPara[0]$HDINT);

//**********************************************************************************************************************************************************
    CMD_SM_GET_MODULE_TYPE:
      pResult^.aData[0]$UDINT := SM_TYPE_SAFETY_MODULE_FSOE;

//**********************************************************************************************************************************************************
    CMD_SM_MODULE_REINIT:
      if b_ReInitMarker then

        // next time we check for the configured state of the cpu
        b_CheckConfigured := TRUE;

        // check again in background
        SetSafetyState(NewState:=_ReinitConfig);

        b_ReInitMarker := FALSE;
      end_if;

//**********************************************************************************************************************************************************
    CMD_SM_POST_INIT_FINISHED:

      // remember that we've been here
      b_PostInitPassed := TRUE;

      Found := FALSE;
      if Online then
        // get configuration if module is configured

        // get state via SDO communication
        sd_retval := SDOStdRequ ( us_Command      := SDO_COMMAND_GET_STATE
                                , p_us_RespData   := ( #GetStateResp )$^USINT
                                , us_RespLength   := sizeof(GetStateResponseType)
                                );

        // the cpu is configured, load the new configuration
        if ( sd_retval = 0 ) &
           (GetStateResp.ConfigState <> CFG_STATE_UNKNOWN) &
           (GetStateResp.ConfigState <> CFG_STATE_INVALID) &
           (GetStateResp.ConfigState <> CFG_STATE_NOT_CONFIGURED) then

          //get configuration from safe CPU and build routing tables
          GetRoutingData();

          Found := TRUE;
        end_if;
      end_if;

      // if we didn't get the config here => try again later
      if Found = FALSE then
        //get configuration from safe CPU and build routing tables later in background
        b_GetNewConfiguration := FALSE;

          // next time we check for the configured state of the cpu
        b_CheckConfigured := TRUE;

        // check again in background
        SetSafetyState(NewState:=_ReinitConfig);
      end_if;

//**********************************************************************************************************************************************************
    CMD_SM_SET_NEW_SYNC_MODE:

//**********************************************************************************************************************************************************
  else
    if bd_LogOnceMarker.InvalidNewInstCmd = FALSE then
      bd_LogOnceMarker.InvalidNewInstCmd := TRUE;
      LogValue("@024A (SafetyBaseFSoE::ClassSvr::NewInst) [SL] Received invalid command: 0x{0}", Value:=pPara^.uiCmd);
    end_if;
//**********************************************************************************************************************************************************
  END_CASE;

END_FUNCTION

FUNCTION VIRTUAL GLOBAL SafetyBaseFSoE::Background
  VAR_INPUT
    EAX 	: UDINT;
  END_VAR
  VAR_OUTPUT
    state (EAX) 	: UDINT;
  END_VAR
  VAR
    sd_retval         : DINT;
    GetStateResp      : GetStateResponseType;
    LastWriteCounter  : UDINT;
    FileHandle        : DINT;
    MyPara 	          : CmdStruct;
    MyResult	        : results;
  END_VAR

  // if any LED is active, then firmware update is not active and we can do our work
  if (VoltageOK | RunState | ServiceMode | ErrorState) then

    // if a quit error is pending
    if QuitComError = 2 then
      MyPara.uiCmd := CMD_SM_QUIT_ERROR_VIA_OS;
      MyPara.aPara[0] := THIS$DINT;
      MyPara.aPara[1] := SafetyNumber$DINT;
      pSafetyManagerThis^.NewInst(#MyPara, #MyResult);

      QuitComError := MyResult.aData[0]$DINT;

      // refresh the server on the outer object
      RefreshAsySrv();
    end_if;

    if (SafetyState = _ReinitConfig) then

      // check every second if the cpu is configured
      if b_CheckConfigured & ((ops.tAbsolute - ud_LastCheckConfig) > 3000) then
        // get state via SDO communication
        sd_retval := SDOStdRequ ( us_Command      := SBF_SDO_COMMAND_GET_STATE
                                , p_us_RespData   := ( #GetStateResp )$^USINT
                                , us_RespLength   := sizeof(GetStateResponseType)
                                );

        // the cpu is configured, load the new configuration
        if ( sd_retval = 0 ) &
           (GetStateResp.ConfigState <> SBF_CFG_STATE_UNKNOWN) &
           (GetStateResp.ConfigState <> SBF_CFG_STATE_INVALID) &
           (GetStateResp.ConfigState <> SBF_CFG_STATE_NOT_CONFIGURED) then

          b_CheckConfigured := FALSE;

          b_GetNewConfiguration := TRUE;
        end_if;

        // remember the last time we checked for configurated cpu
        ud_LastCheckConfig := ops.tAbsolute;
      end_if;

      // if there is a new configuration => get it
      if b_GetNewConfiguration then
        // get configuration from safe CPU and build routing tables
        sd_retval := GetRoutingData();
        if sd_retval = 0 then
          b_GetNewConfiguration := FALSE;

          SendAllUnsafeValues();
        else
          LogError("@024B (SafetyBaseFSoE::Background) FAILED TO REINIT THE SAFECPU: .");
        end_if;
      end_if;
    elsif ConnectionInfos.ConnectionNo then
      // if there are still connections => check if they are initialized
      CheckFSoEConnections();
    end_if;

    // here we save the log file from the module to the harddrive (started by user)
    if DiagVars.SavingLogInProgress then

      case DiagVars.SavingLogSSW of

  // ********************************************************************************************************************************************
        GetLogHeader:     // get log header from module (contains size of log memory and write counter)

          // get log header via SDO communication
          sd_retval := SDORequ ( us_Command      := SBF_SDO_COMMAND_GET_LOG_HDR
                               , p_us_RequData   := #DiagVars.ucChoiceSaveLog
                               , us_RequLength   := 1
                               , p_us_RespData   := ( #DiagVars.LogHeader)$^USINT
                               , us_RespLength   := sizeof(DiagStructType.LogHeader)
                               );

          if ( sd_retval = 0 ) then
            DiagVars.LogMemToGet := DiagVars.LogHeader.LogMemSize;
            DiagVars.pLogFileMem$pVoid := ToStdLib.Malloc(size:=DiagVars.LogHeader.LogMemSize);
            //_memset(dest:=DiagVars.pLogFileMem$pVoid, usByte:=0, cntr:=DiagVars.LogHeader.LogMemSize);
            if DiagVars.ucChoiceSaveLog = 0 then
              DiagVars.ReadBaseAdr := SBF_SDO_ADDRESS_LOG_UC1;
            else
              DiagVars.ReadBaseAdr := SBF_SDO_ADDRESS_LOG_UC2;
            end_if;
            DiagVars.SavingLogSSW := GetLogFileBlocks;

          end_if;

  // ********************************************************************************************************************************************
        GetLogFileBlocks: // get the log memory from the application memory of the module (every cycle only a little bit to prevent runtime error in module)

          // we wait here until UpdateCy finishes our work

  // ********************************************************************************************************************************************
        GetLogHeader2:    // get log header from module again. if write counter changed,
                          // we repeat GetLogFileBlocks. otherwise we continue to save the file

          LastWriteCounter := DiagVars.LogHeader.WriteCounter;

          // get LogHeader
          sd_retval := SDORequ ( us_Command      := SBF_SDO_COMMAND_GET_LOG_HDR
                               , p_us_RequData   := #DiagVars.ucChoiceSaveLog
                               , us_RequLength   := 1
                               , p_us_RespData   := ( #DiagVars.LogHeader)$^USINT
                               , us_RespLength   := sizeof(DiagStructType.LogHeader)
                               );

          if ( sd_retval = 0 ) then

            // if write counter is different, repeat last step
            if DiagVars.LogHeader.WriteCounter <> LastWriteCounter then
              DiagVars.SavingLogSSW := GetLogFileBlocks;

              DiagVars.LogMemToGet := DiagVars.LogHeader.LogMemSize;

              // realloc memory (maybe it's a different size)
              ToStdLib.Free(mptr:=DiagVars.pLogFileMem$pVoid);
              DiagVars.pLogFileMem$pVoid := ToStdLib.Malloc(size:=DiagVars.LogHeader.LogMemSize);
            else
              // write counter is equal. continue to last step
              DiagVars.SavingLogSSW := SaveLogFile;
            end_if;
          end_if;

  // ********************************************************************************************************************************************
        SaveLogFile:      // save the memory to the specified file (DPNE)

          // open file (create/overwrite always)
          FileHandle := FileSys.FileOpen(filename:=#DiagVars.DPNE[0], attributes:=ATT_CREATE_ALWAYS);

          DiagVars.SavingLogSuccessful := 1;

          if FileHandle >= 0 then

            // save content to it
            if FileSys.FileWrite(handle:=FileHandle, buffer:=DiagVars.pLogFileMem, length:=DiagVars.LogHeader.LogMemSize) <> DiagVars.LogHeader.LogMemSize$DINT then
              // failed to write to file
              LogError("@024C (SafetyBaseFSoE::Background) Failed to write to binary LogFile.");
              DiagVars.SavingLogSuccessful := -1;
            end_if;

            // close file
            FileSys.FileClose(handle:=FileHandle);
          else
            // failed to open file
            LogError("@024D (SafetyBaseFSoE::Background) Failed to open binary LogFile.");
            DiagVars.SavingLogSuccessful := -1;
          end_if;

          ToStdLib.Free(mptr:=DiagVars.pLogFileMem$pVoid);
          DiagVars.pLogFileMem := NIL;

          DiagVars.SavingLogSSW := GetLogHeader;
          DiagVars.SavingLogInProgress := FALSE;

      end_case;
    end_if;
  end_if;

  state := READY;

END_FUNCTION

FUNCTION VIRTUAL GLOBAL SafetyBaseFSoE::RtWork
  VAR_INPUT
    EAX 	: UDINT;
  END_VAR
  VAR_OUTPUT
    state (EAX) 	: UDINT;
  END_VAR
  VAR
    calloption    : UDINT;
    PDOLength     : UINT;
    pBuffer       : ^USINT;
    pDOInfo       : ^t_DOInfo;
    i             : USINT;
  END_VAR

  // Save state
  // This must be the 1. line in this function or EAX may be overwritten by the generated AWL code
  calloption := EAX;

  if calloption = CALL_OPTION_RT_PRESCAN then    // Called from UpdateRt

//============================ Profiler start======================================================
#ifdef  DM_Profiler
    StartTimeMeasurement(usMode := DMTIME_RT);
#endif
//============================ Profiler end========================================================

    // do pdo communication only, if module has been found and initialized correctly and if there are some LEDs on (else a FW-Update is running)
    if Online &
       (( SafetyState = _SafetyClassOK ) | ( SafetyState = _WaitForSynchronicity ) | ( SafetyState = _ReinitConfig ) | ( SafetyState = _ModFromCfgNotFound ) | ( SafetyState = _UnknownCfgError ) | ( SafetyState = _UnsafeVarNotFound )) then

      // get I/O state, runstate, error
      UpDateNotStd(calloption:=calloption);

      // wait until the safetymanager has initialized everything
      if b_ManagerInitialisationFinished = FALSE then
        return;
      end_if;

      // if any LED is active, then firmware update is not active and we can do our work
      if (VoltageOK | RunState | ServiceMode | ErrorState) then
        // if we are in run state
        if RunState then
          if PDOSingleRunActive & WriteDOsUsed then
            PDOSingleRunActive -= 1;
            if PDOSingleRunActive = 0 then
              for i := 0 to WriteDOsUsed-1 do
                SetDORunState(Handle:=aWritePDOs[i].Handle, NewState:=_BUS_IF_RUN_STATE_NO_RUN);
              end_for;
            end_if;
          end_if;

          //read PDO from hardware, only if PDO is needed by other moduls
          if ( PDOOutputIsUsed ) & ReadDOsUsed then

            PDOLength := pPDOLengthInfoData^.PDOReadLength;

            // only if length is bigger than minimum and smaller than maximum
            if ( PDOLength >= SBF_SPDO_MIN_LENGTH ) & ( PDOLength <= MyPDOReadSize) then

              pBuffer := #PDOOutputBuffer[0];
              pDOInfo := #aReadPDOs[0];
              for i := 0 to (ReadDOsUsed-1) do
                _memcpy(ptr1:=pBuffer, ptr2:=pDOInfo^.pData, cntr:=pDOInfo^.Length);
                pBuffer += pDOInfo^.Length;
                pDOInfo += sizeof(t_DOInfo);
              end_for;

#ifdef SAFETY_PROTOCOL_ANALYZER_ACTIVATED
  RecordFrame(pFrame:=(#PDOOutputBuffer[0])$^DINT, FrameState:=0, IsFSoEPDO:=TRUE);
#endif
            else
              InvalidPDOSizeCnt += 1;
            end_if;
          end_if;
        end_if;
      end_if;
    end_if;

//============================ Profiler start======================================================
#ifdef  DM_Profiler
    StopTimeMeasurement(usMode := DMTIME_RT);
#endif
//============================ Profiler end========================================================

  elsif calloption = CALL_OPTION_RT_POSTSCAN then // Called from UpdateRtPostScan

//============================ Profiler start======================================================
#ifdef  DM_Profiler
    StartTimeMeasurement(usMode := DMTIME_RTPOSTSCAN);
#endif
//============================ Profiler end========================================================

    // do pdo communication only, if module has been found and initialized correctly and if there are some LEDs on (else a FW-Update is running)
    if Online &
       (( SafetyState = _SafetyClassOK ) | ( SafetyState = _WaitForSynchronicity ) | ( SafetyState = _ModFromCfgNotFound ) | ( SafetyState = _UnknownCfgError ) | ( SafetyState = _UnsafeVarNotFound )) then

      // if any LED is active, then firmware update is not active and we can do our work
      if (VoltageOK | RunState | ServiceMode | ErrorState) then

        // write unsafe I/Os
        UpDateNotStd(calloption:=calloption);

        if RunState & ((us_SetBusReadyState = SetBusReadyFinished) | b_ManualQuit) then
          //write PDO to hardware
          if ( ui_cnt_PDOInputBuffer > 0 ) then
            WritePDO2Module();
          end_if;
        end_if;
      end_if;
    end_if;

//============================ Profiler start======================================================
#ifdef  DM_Profiler
    StopTimeMeasurement(usMode := DMTIME_RTPOSTSCAN);
#endif
//============================ Profiler end========================================================
  end_if;

  state := READY;

END_FUNCTION

FUNCTION VIRTUAL GLOBAL SafetyBaseFSoE::ConnectEvent
  VAR
    MyPara 	              : CmdStruct;
    MyResult	            : results;
  END_VAR

  //start DOs
  StartDO();

  if SafetyState = _ModuleNotFound then
    if ModuleSyncNo = 0 then
      SetSafetyState(NewState:=_SafetyClassOK);
    else
      SetSafetyState(NewState:=_WaitForSynchronicity);
    end_if;
  end_if;

  // if we we're already connected => tell the sdias manager we're back (safetythis has to be valid if b_Reconnect is set, therefore we don't have to check it here)
  if b_Reconnect then
    MyPara.uiCmd := CMD_SM_MODULE_RECONNECT;
    MyPara.aPara[0] := THIS$DINT;
    pSafetyManagerThis^.NewInst(#MyPara, #MyResult);
  end_if;

  // whenever the postinit has passed and we got a connect (module has been plugged in after booting the application) => get it's config
  if b_PostInitPassed = TRUE then
    // start reading the config in background (if we're in init the post-init read-out will be faster)

    // next time we check for the configured state of the cpu
    b_CheckConfigured := TRUE;

    // check again in background
    SetSafetyState(NewState:=_ReinitConfig);
  end_if;

// online is set if module init succeeds
//  Online := 1;

END_FUNCTION

FUNCTION VIRTUAL GLOBAL SafetyBaseFSoE::DisconnectEvent
  VAR
    MyPara 	              : CmdStruct;
    MyResult	            : results;
  END_VAR

  //stop DOs
  StopDO();

  // reset time sync state and tell the manager
  if pSafetyManagerThis then
    MyPara.uiCmd := CMD_SM_MODULE_DISCONNECT;
    MyPara.aPara[0] := THIS$DINT;
    pSafetyManagerThis^.NewInst(#MyPara, #MyResult);

    b_Reconnect := TRUE;
  end_if;

  // clear request, otherwise problems could occur on next connect
  LastRequest := _NoOpenRequest;
  ud_AsyComRetryCounter := 0; // reset retry counter

  SafetyNumber := 0;
  FirmwareVersion := 0;

  // increment the config checksum to ensure the readout on reconnect (config readout also contains check of connected modules)
  DesignerPrjConfigCRC += 1;

  SetSafetyState(NewState:=_ModuleNotFound);

  // remove the cpu from all classes, which use it
  ResetConfig();

  if UnsafeScheduler <> UnsafeSchedulerSetBusReady then
    us_SetBusReadyState := WaitPDOsSyncron;
    UnsafeScheduler := UnsafeSchedulerSetBusReady;
  end_if;

  MaxVarsPerReadPackage := 0;
  ReadFramesNeeded := 0;
  MaxVarsPerWritePackage := 0;
  WriteFramesNeeded := 0;

  Online := 0;

END_FUNCTION

FUNCTION VIRTUAL GLOBAL SafetyBaseFSoE::InterruptEvent

END_FUNCTION

FUNCTION SafetyBaseFSoE::SetDORunState
  VAR_INPUT
    Handle 	: UDINT;
    NewState 	: t_BusIFRunState;
  END_VAR
  VAR
    dataSETRUNSTATE : t_SetRunStateCfg;
    tempCmd : CmdStruct;
    _result : results;
  END_VAR

  // set runstate of read
  dataSETRUNSTATE.Handle      := Handle;
  dataSETRUNSTATE.NewRunState := NewState;

  tempCmd.uiCmd         := _BUS_IF_SET_RUN_STATE;
  tempCmd.aPara[0]      := (#dataSETRUNSTATE)$DINT;

  ToBusInterface.NewInst(pPara:=#tempCmd, pResult:=#_result);

  if _result.aData[0]$t_BusIFRetvalErrorcode <> _BUS_IF_RETVAL_OK then
    if NewState = _BUS_IF_RUN_STATE_NO_RUN then
      DOStopFailCounter += 1;
    else
      DOStartFailCounter += 1;
    end_if;
  end_if;

END_FUNCTION

FUNCTION VIRTUAL GLOBAL SafetyBaseFSoE::CyWork
  VAR_INPUT
    EAX 	: UDINT;
  END_VAR
  VAR_OUTPUT
    state (EAX) 	: UDINT;
  END_VAR
  VAR
    p_SDO_act             : ^SDOHeader;
    us_SDO_length         : USINT;
    i                     : UINT;
    p_ReceiveObj          : pVirtualBase;
    p_SDOviaPath          : ^SDOviaPath;
    sd_retval             : DINT;
    IsStandardResp        : BOOL;
    SDORequestBuffer      : SDORequReadConfig;
    DataLen               : USINT;
    us_UnsafeSchedulerRun : USINT;
    p_PDOInBufferAct      : ^PDOInputBuffer;
    EverythingSynchron    : BOOL;
    MyPara 	              : CmdStruct;
    MyResult	            : results;
    UnsafeWrPackageNo     : USINT;
    aUnsafeWrPackages     : UnsafeWritePackages;
    UnsafeRdPackageNo     : USINT;
    aUnsafeRdPackages     : UnsafeReadPackages;
    TmpVal                : DINT;
    AddUnsafePackage      : BOOL;
    GotNewUnsafeValue     : BOOL;
    pHelpUnsafe           : ^UnsafeIORoutingElement;
    BDINTWriteVars        : USINT;
    pAddDynSlaveResp      : ^t_AddDynSlaveResponse;
  END_VAR

//============================ Profiler start======================================================
#ifdef  DM_Profiler
  StartTimeMeasurement(usMode := DMTIME_CY);
#endif
//============================ Profiler end========================================================

#ifdef HWK_SHOW_PRAGMA_MESSAGES
  if b_LogFirstDone = 1 then
    for i := 0 to (ui_cnt_PDOInputBuffer-1) do
      LogValue("@027F (SafetyBaseFSoE::WritePDO2Module) Copy 0x{0} Bytes to offset 0x{1} of Write PDO Nr. 0x{2}", Value:=aLogValues[i].ByteLen, Value2:=aLogValues[i].Offset, Value3:=aLogValues[i].DOIndex);
    end_for;

    b_LogFirstDone := 2;
  end_if;
#endif

  // do sdo communication only, if module has been found and initialized correctly and if there are some LEDs on (else a FW-Update is running)
  if Online & (VoltageOK | RunState | ServiceMode | ErrorState) &
     (( SafetyState <> _ModuleNotFound ) & ( SafetyState <> _MemAllocFailed ) & ( SafetyState <> _LostPowerSupply ) & ( SafetyState <> _ReadFWVerFailed ) & ( SafetyState <> _WrongSafetyHW )) then

    // wait until the safetymanager has initialized connection
    if (b_ManagerReadyForSDO = FALSE) then
      return;
    end_if;

    //Update of service messages doesn't take place in realtime

    // if we have to quit the communication errors and there is no other request open at this time
    if (QuitComError = 1) & (LastRequest = _NoOpenRequest) then
      if UnsafeScheduler <> UnsafeSchedulerSetBusReady then
        us_SetBusReadyState := WaitPDOsSyncron;
        UnsafeScheduler := UnsafeSchedulerSetBusReady;
      end_if;

      QuitComError := 0;

      // refresh the server on the outer object
      RefreshAsySrv();
    end_if;

    //read SDO from module and send it to the target module
    //check, if SDO is available and valid
    if ( p_Handle_SDO_Read^.us_Status = SAFETY_SDO_DATA_VALID ) then

      //calculate length of SDO
      us_SDO_length := sizeof(SDOHeader.StdHeader.CRC) + p_Handle_SDO_Read^.SDOStructure.SDOHeader.StdHeader.Len;

      //copy SDO without first byte (=status byte)
      ToStdLib.MemCpy(dest := p_SDOOutputBuffer, source := #p_Handle_SDO_Read^.SDOStructure, size := us_SDO_length );

#ifdef SAFETY_PROTOCOL_ANALYZER_ACTIVATED
  RecordFrame(p_SDOOutputBuffer$^DINT, 0);
#endif

      //mark data as received
      p_Handle_SDO_Read^.us_Status := SAFETY_SDO_NO_DATA;

      //find target object for routing
      p_ReceiveObj := NIL;

      IsStandardResp := FALSE;
      //check, if receiver is addressed by safety number or hardware path
      if ((p_SDOOutputBuffer^.SDOHeader.StdHeader.Typ$USINT AND SBF_SSDO_MASK_TYPE)$t_SafetyFrameType = SSDO_MOD) then

        //search this-pointer of receiver with safety number
        p_ReceiveObj := ( GetRoutingPointerByNumber(ud_SafeNumber := p_SDOOutputBuffer^.SDOHeader.DstAdr))$pVirtualBase;

      elsif ((p_SDOOutputBuffer^.SDOHeader.StdHeader.Typ$USINT AND SBF_SSDO_MASK_TYPE)$t_SafetyFrameType = SSDO_MOD_TP) then

        //search this-pointer of receiver with hardware path
        p_SDOviaPath := p_SDOOutputBuffer$^SDOviaPath;
        p_ReceiveObj := ( GetRoutingPointerByPath(p_ActObjectPath := #p_SDOviaPath^.TopologyPath[0], p_SDOviaPath^.StdHeader.Len - 8))$pVirtualBase;
      elsif ((p_SDOOutputBuffer^.SDOHeader.StdHeader.Typ$USINT AND SBF_SSDO_MASK_TYPE)$t_SafetyFrameType = SDO_STD) then
        IsStandardResp := TRUE;
        StandardResponse := (p_SDOOutputBuffer$^StandardFrameType)^;
        if StandardResponse.SDOHeader.SeqNr = (StandardSeqNr OR 16#80) then

          // if the microcontroller got powered again and we have an SDO response => also get the configuration (don't wait the whole time)
          //if b_WaitForFirmwareBoot = TRUE then // no if to be faster (if it's false, it does not matter if we set it again to false)
          b_WaitForFirmwareBoot := FALSE;
          //end_if;

          case LastRequest of
            _NoOpenRequest: // error, no open request, but we got a response
              LogError("@0252 (SafetyBaseFSoE::CyWork) Standard frame response received, without open request.");

            _SetBusReady:
              IF StandardResponse.SDOHeader.Cmd = SBF_SDO_COMMAND_SET_BUS_READY THEN
                if us_SetBusReadyState <> SendSetBusReady then
                  LogError("@0253 (SafetyBaseFSoE::CyWork) Got Response of SetBusReady, but SSW is not in the right step.");
                  return;
                end_if;
                us_SetBusReadyState := SetBusReadyFinished;
                b_ManualQuit := FALSE;
                UnsafeScheduler := UnsafeSchedulerGetDiagVars; // Go on with the action-steps, done here so we don't lose a whole cycle
                LastRequest := _NoOpenRequest;
                ud_AsyComRetryCounter := 0; // reset retry counter
                if SafetyState = _WaitForSynchronicity then
                  SetSafetyState(NewState:=_SafetyClassOK);
                end_if;
              else
                LogError("@0256 (SafetyBaseFSoE::CyWork) Invalid command: bus ready expected.");
              END_IF;

            _ReadData:
              // if we did read command, then save the value to corresponding server
              if StandardResponse.SDOHeader.Cmd = SBF_SDO_COMMAND_READ then
                // if returncode is 0 read succeeded
                if StandardResponse.aData[0] = 0 then
                  // check if length is correct
                  if StandardResponse.aData[1] = StandardRequest.aData[4] then
                    // delete request
                    LastRequest := _NoOpenRequest;
                    ud_AsyComRetryCounter := 0; // reset retry counter

                    if (DiagVars.SavingLogSSW = GetLogFileBlocks) then
                      // save the last block in the memory for the file
                      _memcpy(ptr1:=DiagVars.pLogFileMem$pVoid + (DiagVars.LogHeader.LogMemSize - DiagVars.LogMemToGet),
                              ptr2:=#StandardResponse.aData[2],
                              cntr:=DiagVars.BytesToGet);

                      DiagVars.LogMemToGet -= DiagVars.BytesToGet;

                      if DiagVars.LogMemToGet = 0 then
                        DiagVars.SavingLogSSW := GetLogHeader2;
                      end_if;
                    else
                      LogError("@0255 (SafetyBaseFSoE::CyWork) SDO Receive: Invalid Read response (no diagnostic read active).");
                    end_if;
                  end_if;
                end_if;
              else
                LogError("@0256 (SafetyBaseFSoE::CyWork) SDO Receive: Invalid command, read expected.");
              end_if;

            _ReadValues:
              // if we did read command, then save the value to corresponding server
              if StandardResponse.SDOHeader.Cmd = SBF_SDO_COMMAND_READ_VALUES then
                // if returncode is 0 read succeeded
                if StandardResponse.aData[0] = 0 then
                  // check if length is correct
                  if StandardResponse.aData[1] = StandardRequest.aData[0] then
                    // delete request
                    LastRequest := _NoOpenRequest;
                    ud_AsyComRetryCounter := 0; // reset retry counter

                    // if we got some outputs in the routing table and a valid pointer, write values to servers
                    if ui_CntUnsafeOutputs & pUnsafeOutElement then

                      // depending on length we do different number of server write-methods to set the data we just read
//                      pUnsafeOutElement := p_UnsafeOutputsTable + (UnsafeReadTransNr * MaxVarsPerReadPackage * sizeof(UnsafeIORoutingElement));  // the pointer is already on this element
                      for i := 0 to (StandardResponse.aData[1] - 1) do
                        // save the new value temporarily
                        TmpVal := StandardResponse.aData[2 + (i * sizeof(DINT))]$DINT;
                        if pUnsafeOutElement^.ud_Thisp then
                          if pUnsafeOutElement^.UnsafeType = BDINTOutput then
                            pUnsafeOutElement^.sd_OldValue := RD(pUnsafeOutElement^.ud_Thisp$^void)$DINT;
                            TmpVal := ((pUnsafeOutElement^.sd_OldValue$UDINT AND (NOT pUnsafeOutElement^.BitMask)) OR
                                      (TmpVal$UDINT AND pUnsafeOutElement^.BitMask))$DINT;

                            // now we have to write the value to the server
                            WR(pUnsafeOutElement^.ud_Thisp$^void, TmpVal);
                          else
                            WR(pUnsafeOutElement^.ud_Thisp$^void, TmpVal);
                          end_if;
                        elsif (pUnsafeOutElement^.UnsafeType = ExternalOutput) | (pUnsafeOutElement^.UnsafeType = ExternalBDINTOutput) then
                          pUnsafeOutElement^.sd_NewValue4External := TmpVal;

                          // mark the value as valid
                          pUnsafeOutElement^.b_IsValid := TRUE;
                        end_if;
                        pUnsafeOutElement += sizeof(UnsafeIORoutingElement);
                      end_for;
                    end_if;

                    UnsafeReadTransNr += 1;
                  end_if;
                end_if;
              else
                LogError("@0257 (SafetyBaseFSoE::CyWork) SDO Receive: Invalid command, read values expected.");
              end_if;

            _WriteValues:
              if IsOptimizedCPU() then
                // if we did a write command, just check
                if StandardResponse.SDOHeader.Cmd = SBF_SDO_COMMAND_WRITE_VALUES then
                  // delete request
                  LastRequest := _NoOpenRequest;
                  ud_AsyComRetryCounter := 0; // reset retry counter

                  // if there is no more element to send or check for changes => proceed to the next step
                  if pUnsafeInElement = NIL then
                    UnsafeScheduler := UnsafeSchedulerReadData; //We need to set scheduler to next step....
                  end_if;
                else
                  LogError("@0258 (SafetyBaseFSoE::CyWork) SDO Receive: Invalid command, write expected.");
                end_if;
              else
                // on CSCP011 the SDO_COMMAND_WRITE_VALUES didn't exist

                // if we did a write command, just check
                if StandardResponse.SDOHeader.Cmd = SBF_SDO_COMMAND_WRITE then
                  // delete request
                  LastRequest := _NoOpenRequest;
                  ud_AsyComRetryCounter := 0; // reset retry counter

                  if UnsafeWriteTransNr < (WriteFramesNeeded - 1) then
                    UnsafeWriteTransNr += 1;
                  else
                    UnsafeWriteTransNr := 0;
                    UnsafeWritingActive := FALSE;
                    UnsafeScheduler := UnsafeSchedulerReadData; //We need to set scheduler to next step....
                  end_if;
                else
                  LogError("@0258 (SafetyBaseFSoE::CyWork) SDO Receive: Invalid command, write expected.");
                end_if;
              end_if;

            _GetCRC:
              // check if it's a response to a read command
              if StandardResponse.SDOHeader.Cmd = SBF_SDO_COMMAND_READ then
                // if returncode is 0 read succeeded
                if StandardResponse.aData[0] = 0 then
                  // check if length is correct
                  if StandardResponse.aData[1] = 4 then

                    // delete request
                    LastRequest := _NoOpenRequest;
                    ud_AsyComRetryCounter := 0; // reset retry counter

                    if DesignerPrjConfigCRC <> StandardResponse.aData[2]$UDINT then
                      // CRC has changed => save the new crc
                      DesignerPrjConfigCRC := StandardResponse.aData[2]$UDINT;

                      // show that we read the config of the class again
                      SetSafetyState(NewState:=_ReinitConfig);

                      if pSafetyManagerThis then
                        MyPara.uiCmd := CMD_SM_NEW_SAFETY_PROJECT;
                        MyPara.aPara[0] := 4;
                        MyPara.aPara[4] := (#SafetyNumber)$DINT;
                        pSafetyManagerThis^.NewInst(#MyPara, #MyResult);
                      end_if;

                      // remove the cpu from all classes, which use it
                      ResetConfig();

                      // we have to return here because:
                      // the command CMD_SM_NEW_SAFETY_PROJECT will trigger a disconnect of this class which will set the unsafe scheduler to setbusready,
                      // which would skip the synchron check in the actual cyclic run because everything of the old configuration is synchron now
                      return;
                    end_if;
                  end_if;
                end_if;
              end_if;

            _WriteSysTime:
              if StandardResponse.SDOHeader.Cmd = SBF_SDO_COMMAND_WRITE then
                // if returncode is 0 read succeeded
                if StandardResponse.aData[0] = 0 then
                  // delete request
                  LastRequest := _NoOpenRequest;
                  ud_AsyComRetryCounter := 0; // reset retry counter
                end_if;
              else
                LogError("@0258 (SafetyBaseFSoE::CyWork) SDO Receive: Invalid command, write expected.");
              end_if;

            _WriteFlexConCommand:
              if StandardResponse.SDOHeader.Cmd = SBF_SDO_COMMAND_WRITE then
                // if returncode is 0 read succeeded
                if StandardResponse.aData[0] = 0 then
                  // delete request
                  LastRequest := _NoOpenRequest;
                  ud_AsyComRetryCounter := 0; // reset retry counter
                end_if;
              else
                LogError("@0258 (SafetyBaseFSoE::CyWork) SDO Receive: Invalid command, write expected.");
              end_if;

            _DiagState:
              if StandardResponse.SDOHeader.Cmd = SBF_SDO_COMMAND_GET_STATE then
                _memcpy(ptr1 := #DiagVars.UserGetStateResp,
                        ptr2 := #StandardResponse.aData + SIZEOF(USINT),
                        cntr := sizeof(GetStateResponseType) );
                DiagVars.UserDiagStateReady := TRUE;
                DiagVars.UserWantsDiagState := FALSE;
                LastRequest := _NoOpenRequest;
                ud_AsyComRetryCounter := 0; // reset retry counter
              end_if;
            _DiagInfo:
              if StandardResponse.SDOHeader.Cmd = SBF_SDO_COMMAND_GET_DIAG_INFO then
                _memcpy(ptr1 := #DiagVars.UserGetDiagInfoResp,
                        ptr2 := #StandardResponse.aData + SIZEOF(USINT),
                        cntr := sizeof(SafetyDiagInfo) );
                DiagVars.UserDiagInfoReady := TRUE;
                DiagVars.UserWantsDiagInfo := FALSE;
                LastRequest := _NoOpenRequest;
                ud_AsyComRetryCounter := 0; // reset retry counter
              end_if;

            _ReadRetryCounter:
              //if we did read command, then save the value to corresponding server
              if StandardResponse.SDOHeader.Cmd = SBF_SDO_COMMAND_READ then
                // if returncode is 0 read succeeded
                if StandardResponse.aData[0] = 0 then
                  // check if length is correct
                  if StandardResponse.aData[1] = SBF_SDO_LENGTH_RETRY_COUNTER then
                    // delete request
                    LastRequest := _NoOpenRequest;
                    ud_AsyComRetryCounter := 0; // reset retry counter

                    //Only Write if Retry Counter has changed
                    if StandardResponse.aData[2] <> us_OldRetryCounter then
                      //if retry counter has changed, save the new retry counter
                      SafetyRetryCounter += to_usint(StandardResponse.aData[2] - us_OldRetryCounter);
                      us_OldRetryCounter := StandardResponse.aData[2];

                      //0x20400000 is adress of retry counter: 1 byte amount of all retries of all modules, 16byte µC1, 16 byte µC2
                      //Save the values from the modules
                      ToStdLib.MemCpy(dest:=#a_RetryCnt[0], source:=#StandardResponse.aData[3], size:=SBF_SDO_LENGTH_RETRY_COUNTER);

                      //Calls the method of class sdiassafetymanager
                      SetRetryCounter();
                    end_if;
                  end_if;
                end_if;
              else
                LogError("@0257 (SafetyBaseFSoE::CyWork) SDO Receive: Invalid command, read values expected.");
              end_if;

            _ErrorChannelInfo:
              //if we did read command, then save the value to corresponding server
              if StandardResponse.SDOHeader.Cmd = SBF_SDO_COMMAND_READ then
                // if returncode is 0 read succeeded
                if StandardResponse.aData[0] = 0 then
                  // check if length is correct
                  if StandardResponse.aData[1] <> 0  then
                    _memcpy(ptr1 := #aErrorMem[actoffset],
                            ptr2 := #StandardResponse.aData[2],
                            cntr := StandardResponse.aData[1]);
                    if remainingPacketlength = 0 then
                      remainingPacketlength := StandardResponse.aData[2] - StandardResponse.aData[1];
                      actoffset := StandardResponse.aData[1];
                    else
                      remainingPacketlength -= StandardResponse.aData[1];
                      actoffset += StandardResponse.aData[1];
                    end_if;

                    // delete request
                    LastRequest := _NoOpenRequest;
                    ud_AsyComRetryCounter := 0; // reset retry counter
                    if remainingPacketlength <= 0  then
                      //Finish
                      DiagVars.UserErrorInfoReady := TRUE;
                      DiagVars.UserWantsErrorInfo := FALSE;
                      remainingPacketlength := 0; //reset remainingPacketlength
                      actoffset := 0; //reset offset
                    end_if;
                  end_if;
                end_if;
              end_if;

            _ReadFlexConNodeState:
              //if we did read command, then save the value to corresponding server
              if StandardResponse.SDOHeader.Cmd = SBF_SDO_COMMAND_READ then
                // if returncode is 0 read succeeded
                if StandardResponse.aData[0] = 0 then
                  // check if length is correct
                  if StandardResponse.aData[1] = sizeof(t_FlexConNodeState) then

                    // store the structure locally
                    _memcpy(ptr1 := #sFlexCon.LastNodeState,
                            ptr2 := #StandardResponse.aData[2],
                            cntr := StandardResponse.aData[1]);

                    // save the values to the server of the object
                    sFlexCon.pCommand^            := sFlexCon.LastNodeState.Command;
                    sFlexCon.pStateMachine^       := sFlexCon.LastNodeState.StateMachine;
                    sFlexCon.pHostSafetyNumber^   := sFlexCon.LastNodeState.HostSafetyNumber;

                    // delete request
                    LastRequest := _NoOpenRequest;
                    ud_AsyComRetryCounter := 0; // reset retry counter
                  end_if;
                end_if;
              end_if;

            _ReadFlexConHostState:
              //if we did read command, then save the value to corresponding server
              if StandardResponse.SDOHeader.Cmd = SBF_SDO_COMMAND_READ then
                // if returncode is 0 read succeeded
                if StandardResponse.aData[0] = 0 then
                  // check if length is correct (maximum the requested size)
                  if StandardResponse.aData[1] & (StandardResponse.aData[1] <= sFlexCon.LastHostState.LastRequestedLength) then
                    // if the size in the response is smaller than the requested (we already got everything in the first package)
                    if StandardResponse.aData[1] <= sFlexCon.LastHostState.LastRequestedLength then
                      // adjust the last requested length to the received for correct handling of the received data
                      sFlexCon.LastHostState.LastRequestedLength := StandardResponse.aData[1];
                    end_if;

                    // if it's the first package
                    if sFlexCon.LastHostState.CurrentReadOffset = 0 then
                      // if length is ok and there is at least 1 connection but not more than the maximum
                      if (StandardResponse.aData[1] >= sizeof(HDINT)) & StandardResponse.aData[2]$HDINT & (StandardResponse.aData[2]$HDINT <= MAX_FSOE_CONNECTIONS) then
                        // the first 4 byte contain the number of connections following
                        sFlexCon.LastHostState.NoConnections := StandardResponse.aData[2]$HDINT;
                        _memcpy(ptr1:=#sFlexCon.LastHostState.aConnections[0], ptr2:=#StandardResponse.aData[2] + sizeof(HDINT), cntr:=sFlexCon.LastHostState.LastRequestedLength - sizeof(HDINT));

                        // calculate how many bytes are missing (what do we need minus what do we already have)
                        sFlexCon.LastHostState.BytesMissing       := sFlexCon.LastHostState.NoConnections$UINT * sizeof(HDINT) + sizeof(HDINT) - sFlexCon.LastHostState.LastRequestedLength;
                        sFlexCon.LastHostState.CurrentReadOffset  += sFlexCon.LastHostState.LastRequestedLength;
                      else
                        // no connection or too many to fit into the array
                        sFlexCon.LastHostState.NoConnections := 0;

                        // nothing missing
                        sFlexCon.LastHostState.BytesMissing := 0;
                      end_if;
                    else
                      // offset is not zero => follow up package
                      _memcpy(ptr1:=#sFlexCon.LastHostState.aConnections[0] + sFlexCon.LastHostState.CurrentReadOffset - sizeof(HDINT), ptr2:=#StandardResponse.aData[2], cntr:=sFlexCon.LastHostState.LastRequestedLength);

                      // update the bytes missing and the current reading offset
                      sFlexCon.LastHostState.BytesMissing      -= sFlexCon.LastHostState.LastRequestedLength;
                      sFlexCon.LastHostState.CurrentReadOffset += sFlexCon.LastHostState.LastRequestedLength;
                    end_if;
                  else
                    // wrong length => reset number of connections
                    sFlexCon.LastHostState.NoConnections := 0;

                    // nothing missing
                    sFlexCon.LastHostState.BytesMissing := 0;
                  end_if;

                  // if we got all data
                  if sFlexCon.LastHostState.BytesMissing = 0 then

                    // update connection state at managing modules
                    MyPara.uiCmd := CMD_SM_UPDATE_FLEX_CON_HOST;
                    MyPara.aPara[0] := sFlexCon.LastHostState.NoConnections$DINT;
                    MyPara.aPara[1] := (#sFlexCon.LastHostState.aConnections[0])$DINT;
                    pSafetyManagerThis^.NewInst(#MyPara, #MyResult);

                    // reset the offset so we start reading at 0 in the next round
                    sFlexCon.LastHostState.CurrentReadOffset := 0;

                    // reset timemark
                    sFlexCon.ud_LastHostStateTimeStamp := ops.tAbsolute;
                  end_if;

                  // delete request
                  LastRequest := _NoOpenRequest;
                  ud_AsyComRetryCounter := 0; // reset retry counter

                end_if;
              end_if;

          else
            LogError("@025A (SafetyBaseFSoE::CyWork) SDO Receive: Invalid standard frame response.");
          end_case;

          // if request is deleted, increase sequence number to set next request
          if LastRequest = _NoOpenRequest then
            if StandardSeqNr < 16#7F then
              StandardSeqNr += 1;
            else
              StandardSeqNr := 0;
            end_if;
          end_if;
        else
          LogError("@025B (SafetyBaseFSoE::CyWork) SDO Receive: Invalid sequence number in Standard SDO response.");
          LogValue("expected: 0x{0} / received: 0x{1}", Value:=(StandardSeqNr OR 16#80), Value2:=StandardResponse.SDOHeader.SeqNr);
        end_if;
      elsif ((p_SDOOutputBuffer^.SDOHeader.StdHeader.Typ$USINT AND SBF_SSDO_MASK_TYPE)$t_SafetyFrameType = SSDO_MOD_DEVADDR) then

        //Check if we know our target
        p_ReceiveObj := ( GetRoutingPointerByNumber(ud_SafeNumber := p_SDOOutputBuffer^.SDOHeader.DstAdr))$pVirtualBase;

        //Forward data to manager if we found no routing target, otherwise the SDO will be directly send to target
        if p_ReceiveObj = NIL then

          // Forward to manager if possible
          if pSafetyManagerThis & us_SDO_length then
  #ifdef DO_DEBUG
            DOCheck(pFrame:=(p_SDOOutputBuffer)$^t_SDOStdHeader, pCheckStruct:=#SDORead);
  #endif

            if ( (p_SDOOutputBuffer^.SDOHeader.StdHeader.Cmd = SBF_SDO_COMMAND_ADD_DYN_SLAVE) | (p_SDOOutputBuffer^.SDOHeader.StdHeader.Cmd = SBF_SDO_COMMAND_ADD_DYN_SLAVE2) )&
               (p_SDOOutputBuffer^.SDOHeader.StdHeader.Typ$USINT AND SBF_SSDO_MASK_RESPONSE) then
              // we need a response big enough to hold our info, the returncode must be 0 and the offset/length info has to be plausible
              if ((p_SDOOutputBuffer^.SDOHeader.StdHeader.Len + sizeof(SDOHeader.StdHeader.CRC)) >= sizeof(t_AddDynSlaveResponse)) &
                  (p_SDOOutputBuffer^.us_Returncode = 0) & CheckAddDynSlaveResponse(p_SDOOutputBuffer$^t_AddDynSlaveResponse) then

                pAddDynSlaveResp := p_SDOOutputBuffer$^t_AddDynSlaveResponse;

                MyPara.aPara[2]       := THIS$DINT;

                MyPara.aPara[3]$HDINT := pAddDynSlaveResp^.OffsetSafeOutData; // offset to data from module
                MyPara.aPara[4]$HDINT := pAddDynSlaveResp^.LenSafeOutData;    // size of data from module

                MyPara.aPara[5]$HDINT := pAddDynSlaveResp^.OffsetSafeInData;  // offset to data to module
                MyPara.aPara[6]$HDINT := pAddDynSlaveResp^.LenSafeInData;     // size of data to module
              else
                _memset(dest:=#MyPara.aPara[2], usByte:=0, cntr:=5*sizeof(DINT));
              end_if;
            end_if;

            MyPara.uiCmd := CMD_SM_SDO_TO_MANAGER;
            MyPara.aPara[0] := to_dint(us_SDO_length);
            MyPara.aPara[1] := p_SDOOutputBuffer$DINT;
            pSafetyManagerThis^.NewInst(#MyPara, #MyResult);

            IsStandardResp := TRUE;
          else
            //log not routable SDOs
            LogValue("@025E (SafetyBaseFSoE::CyWork) Safety module 0x{0}: SDO not routed to receiver {1}", SafetyNumber$UDINT, p_SDOOutputBuffer^.SDOHeader.DstAdr$UDINT);
          end_if;
        end_if;
      else
        LogError("@025C (SafetyBaseFSoE::CyWork) SDO Receive: Invalid frametype in Standard SDO response.");
      end_if;

      //if there is no object, the message will be lost
      if ( p_ReceiveObj ) then

        //send SDO to receiver object
        MyPara.uiCmd := CMD_SM_ADD_SDO_TO_BUFFER;
        MyPara.aPara[0] := p_SDOOutputBuffer$DINT;
        MyPara.aPara[1] := us_SDO_length;
        sd_retval$iprStates := p_ReceiveObj^.NewInst(#MyPara, #MyResult);

//        sd_retval := p_ReceiveObj^.AddSDOToBuffer(p_us_Message := p_SDOOutputBuffer$^USINT, us_length := us_SDO_length);

        if sd_retval$iprStates = ERROR then
          // generate error message with returncode (add to logfile and debugger trace)
          LogValue("@025D (SafetyBaseFSoE::CyWork) AddSDOToBuffer failed: Returncode: -0x{0}", Value:=(0-sd_retval)$UDINT);
        end_if;

      elsif IsStandardResp = FALSE then

        if pSafetyManagerThis & us_SDO_length then
#ifdef DO_DEBUG
          DOCheck(pFrame:=(p_SDOOutputBuffer)$^t_SDOStdHeader, pCheckStruct:=#SDORead);
#endif

          // if the command is get safety number and the compressed path type is 2, it can only be in this system (no interface frame) and therefore forwarding to the manager would not make sense (the class should already find the other module with GetRoutingPointerByPath()
          if (p_SDOOutputBuffer^.SDOHeader.StdHeader.Cmd = SBF_SDO_COMMAND_GET_SAFENBR) &
             (p_SDOOutputBuffer^.SDOHeader.StdHeader.Typ = SSDO_MOD_TP) &
             (p_SDOOutputBuffer^.SDOHeader.DstAdr$USINT = 2) then
            // skip forwarding in this case
          else
            // forward it to the safety manager
            MyPara.uiCmd := CMD_SM_SDO_TO_MANAGER;
            MyPara.aPara[0] := to_dint(us_SDO_length);
            MyPara.aPara[1] := p_SDOOutputBuffer$DINT;
            pSafetyManagerThis^.NewInst(#MyPara, #MyResult);
          end_if;
        else
          //log not routable SDOs
          LogValue("@025E (SafetyBaseFSoE::CyWork) Safety module 0x{0}: SDO not routed to receiver {1}", SafetyNumber$UDINT, p_SDOOutputBuffer^.SDOHeader.DstAdr$UDINT);
        end_if;
      end_if;

    elsif (LastRequest <> _NoOpenRequest) & (ud_TransfertimePerPackage > 0) then
      // count up for timeout
      ud_UnsafeTimeoutCounter += 1;

      if ( ud_UnsafeTimeoutCounter ) > ( 50 * ud_TransfertimePerPackage ) then
        CASE UnsafeScheduler OF

          UnsafeSchedulerSetBusReady:
            LogError("@025F (SafetyBaseFSoE::UpdateCy) Timeout on setting bus ready.");

          UnsafeSchedulerGetDiagVars:
            IF LastRequest = _ReadData THEN
              LogError("@0260 (SafetyBaseFSoE::UpdateCy) Timeout requesting DiagVars.");
            END_IF;
            UnsafeScheduler := UnsafeSchedulerNonPriorData;
            DiagVars.SavingLogSSW := GetLogFileBlocks;

          UnsafeSchedulerNonPriorData:
            if LastRequest = _WriteSysTime then
              LogError("@0497 (SafetyBaseFSoE::UpdateCy) Timeout writing the system time to module.");
            else
              LogError("@0261 (SafetyBaseFSoE::UpdateCy) Timeout requesting CRC.");
            end_if;

            UnsafeScheduler := UnsafeSchedulerWriteData;

          UnsafeSchedulerWriteData:
            LogError("@0262 (SafetyBaseFSoE::UpdateCy) Timeout writing Data 'Unsafe Input'.");
            UnsafeScheduler := UnsafeSchedulerReadData;
            UnsafeWriteTransNr := 0;

          UnsafeSchedulerReadData:
            LogError("@0263 (SafetyBaseFSoE::UpdateCy) Timeout reading Data 'Unsafe Output'.");
            UnsafeScheduler := UnsafeSchedulerDiagState;
            UnsafeReadTransNr := 0;

          UnsafeSchedulerDiagState:
            LogError("@0264 (SafetyBaseFSoE::UpdateCy) Timeout on reading DiagState.");
            UnsafeScheduler := UnsafeSchedulerDiagInfo;

          UnsafeSchedulerDiagInfo:
            LogError("@0265 (SafetyBaseFSoE::UpdateCy) Timeout on reading DiagInfo.");
            UnsafeScheduler := UnsafeSchedulerGetRetryCounter;

          UnsafeSchedulerGetRetryCounter:
            LogError("@0266 (SafetyBaseFSoE::UpdateCy) Timeout on reading RetryCounter.");
            UnsafeScheduler := UnsafeSchedulerChannelError;

          UnsafeSchedulerChannelError:
            LogError("@0267 (SafetyBaseFSoE::UpdateCy) Timeout on reading ChannelErrorInfo.");
            UnsafeScheduler := UnsafeSchedulerGetFlexConNodeState;

          UnsafeSchedulerGetFlexConNodeState:
            LogError("@0267 (SafetyBaseFSoE::UpdateCy) Timeout on reading FlexConNodeState.");
            UnsafeScheduler := UnsafeSchedulerGetFlexConHostState;

          UnsafeSchedulerGetFlexConHostState:
            LogError("@0267 (SafetyBaseFSoE::UpdateCy) Timeout on reading FlexConHostState.");
            UnsafeScheduler := UnsafeSchedulerGetDiagVars;

        END_CASE;

        // we only increase the retry counter if the module is running
        if RunState then
          ud_AsyComRetryCounter += 1;
        end_if;

        if ud_AsyComRetryCounter >= SBF_SDO_MAX_TRIES then
          SetSafetyState(NewState:=_AsyncComError);
          LogError("@0268 (SafetyBaseFSoE::UpdateCy) Too many consecutive asynchronous commands failed! Please contact Sigmatek Support!");
        else
          LastRequest := _NoOpenRequest;
          // if request is deleted, increase sequence number to set next request
          if StandardSeqNr < 16#7F then
            StandardSeqNr += 1;
          else
            StandardSeqNr := 0;
          end_if;
        end_if;
      end_if;
